FUNCTION_BLOCK logiBUS_QD_DIMMER_G (* Dimmer like in the living room for lamps and LEDs, with gamma correction, on a 13-bit PWM output *)
  (* Description: Copyright (c) 2026 HR Agrartechnik GmbH This program and the accompanying materials are made available under the terms of the Eclipse Public License 2.0 which is available at https://www.eclipse.org/legal/epl-2.0/ SPDX-License-Identifier: EPL-2.0 *)
  (* Version 1.0, 2026-11-07, Franz Höpfinger, HR Agrartechnik GmbH, initial version, gamma variant of logiBUS_QD_DIMMER *)
  PACKAGE logiBUS::io::DQ;
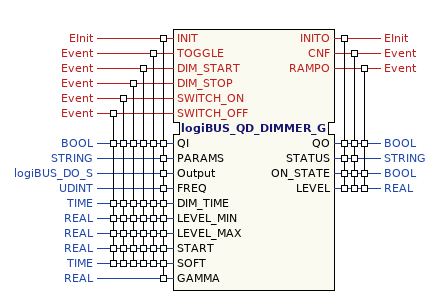
  EVENT_INPUT
    INIT : EInit WITH QI, PARAMS, Output, FREQ, DIM_TIME, LEVEL_MIN, LEVEL_MAX, START, SOFT, GAMMA; (* Service Initialization *)
    TOGGLE WITH QI, DIM_TIME, LEVEL_MIN, LEVEL_MAX, START, SOFT; (* Short press (BUTTON_SINGLE_CLICK of logiBUS_IE): off -> on with the stored brightness (first time START), on -> off; ramp time SOFT *)
    DIM_START WITH QI, DIM_TIME, LEVEL_MIN, LEVEL_MAX, START, SOFT; (* Long press begins (BUTTON_LONG_PRESS_START): dim stepless towards LEVEL_MAX or LEVEL_MIN. Every long press changes the direction, the first one after switching on dims down; at the end it dims the other way. From off: on and dim up *)
    DIM_STOP WITH QI, DIM_TIME, LEVEL_MIN, LEVEL_MAX, START, SOFT; (* Long press ends (BUTTON_LONG_PRESS_UP): stop dimming, the brightness stays and is stored *)
    SWITCH_ON WITH QI, DIM_TIME, LEVEL_MIN, LEVEL_MAX, START, SOFT; (* Switch on directly with the stored brightness (nothing happens if already on) *)
    SWITCH_OFF WITH QI, DIM_TIME, LEVEL_MIN, LEVEL_MAX, START, SOFT; (* Switch off directly, e.g. central off (nothing happens if already off) *)
  END_EVENT
  EVENT_OUTPUT
    INITO : EInit WITH QO, STATUS, ON_STATE, LEVEL; (* Initialization Confirm *)
    CNF WITH QO, STATUS, ON_STATE, LEVEL; (* Confirmation of TOGGLE, DIM_START, DIM_STOP, SWITCH_ON, SWITCH_OFF *)
    RAMPO WITH QO, ON_STATE, LEVEL; (* Ramp finished: LEVEL_MIN or LEVEL_MAX reached while dimming, or switching on/off finished. Not after DIM_STOP *)
  END_EVENT
  VAR_INPUT
    QI : BOOL; (* Event Input Qualifier *)
    PARAMS : STRING; (* Service Parameters *)
    Output : logiBUS::io::DQ::logiBUS_DO_S := logiBUS_DO::Invalid; (* Identify the Output Output_Q1..Q8 *)
    FREQ : UDINT := 400; (* PWM frequency in Hz, read at INIT. Outputs with the same frequency share an LEDC timer (4 timers, LED blinking uses one). Power stage limits, not checked: APIXON 15 PWR Q1 (BTH50030) max. 100 Hz; BTS7030/BTT6030/BTH6070 for valves 100..200 Hz; Trainer20 without power stage *)
    DIM_TIME : TIME := T#4s; (* Time for the whole range LEVEL_MIN..LEVEL_MAX while dimming; a shorter rest takes proportionally less time, so the speed is always the same *)
    LEVEL_MIN : REAL := 10.0; (* Lowest brightness for dimming in % (0..100) *)
    LEVEL_MAX : REAL := 100.0; (* Highest brightness for dimming in % (0..100) *)
    START : REAL := 100.0; (* Brightness in % for the first switching on, before anything is stored *)
    SOFT : TIME := T#300ms; (* Ramp time for switching on and off (TOGGLE, SWITCH_ON, SWITCH_OFF). T#0ms = jump *)
    GAMMA : REAL := 2.2; (* Gamma of the brightness curve, read at INIT: duty = 8191 * (brightness / 8191)^GAMMA. 1.0 = linear (like logiBUS_QD_DIMMER), 2.2 = sRGB (default), 2.6 / 2.8 = Espressif examples, often more even on LEDs. Invalid values (<= 0, not finite) run linear like 1.0 *)
  END_VAR
  VAR_OUTPUT
    QO : BOOL; (* Event Output Qualifier *)
    STATUS : STRING; (* Service Status *)
    ON_STATE : BOOL; (* TRUE = on, FALSE as soon as switching off begins *)
    LEVEL : REAL; (* Brightness in %: on CNF the target of switching on/off or the stopped brightness, on RAMPO the brightness reached *)
  END_VAR
END_FUNCTION_BLOCK
